Fanuc KAREL source: kx00027.KL

-- PROVISIONAL review KL for V1013-1; original PC SHA256 9b216a07d614e4f6a598633b79820f5f10cdf907254fc4f3a3c8d4242918e261
-- Incomplete behavior may be omitted. Consult companion uncertainty JSON. Do not deploy.
PROGRAM KX00027
%NOLOCKGROUP
VAR
  I : INTEGER
  J : INTEGER
  B : BOOLEAN
  F : FILE
  S : STRING[80]
-- UNRESOLVED_DECL P type=000102
BEGIN
  -- UNRESOLVED_PC offsets 5-12; opcodes 9D,23
  -- UNRESOLVED_PC offsets 17-21; opcodes 7F
END KX00027
